(* IEC 61131-3 sources: bevling_machine/framework/sources/04_Machine, 9 files *)

(* ---- F_RecipeValid.st ---- *)
(* 模块说明：检查框架允许的料型、速度、行程和位置顺序。通过仅表示符合示例边界，不代表实机参数已经确认。 *)
FUNCTION F_RecipeValid : BOOL
VAR_INPUT
    stRecipe : ST_Recipe; (* 待校验配方或上层传入的运行配方，字段含义见 ST_Recipe。 *)
END_VAR
FUNCTION F_RecipeValid : BOOL
(* 示例边界：切长 0..1200、速度 0..300、角度正负360，并要求机械手回位<后退<前进<拉料。边界是否适合实机仍需标定。 *)
(* 料型只认 300/450/600：现场侧挡是三个固定位置的气缸，没有 400 这个档；400 是早期仿真的占位值。 *)
F_RecipeValid := ((stRecipe.uiMaterialModel = 300) OR
    (stRecipe.uiMaterialModel = 450) OR (stRecipe.uiMaterialModel = 600))
    AND (stRecipe.lrCutLength > 0.0) AND (stRecipe.lrCutLength <= 1200.0)
    AND (stRecipe.lrCutVelocity > 0.0) AND (stRecipe.lrCutVelocity <= 300.0)
    AND (stRecipe.lrReturnVelocity > 0.0) AND (stRecipe.lrReturnVelocity <= 300.0)
    AND (stRecipe.lrPositionVelocity > 0.0) AND (stRecipe.lrPositionVelocity <= 100.0)
    AND (stRecipe.lrBeltVelocity > 0.0) AND (stRecipe.lrBeltVelocity <= 100.0)
    AND (stRecipe.lrSpindleVelocity > 0.0) AND (stRecipe.lrSpindleVelocity <= 100.0)
    AND (stRecipe.tStepTimeout >= T#1S) AND (stRecipe.tCutTimeout >= T#1S) AND (stRecipe.tSpray > T#0MS)
    AND (ABS(stRecipe.lrCutHome) <= 500.0)
    (* 终点 = 回刀起点 + 切割行程；行程放到 1200 后，终点上限相应放到 1300（典型 100+1200）。 *)
    AND (ABS(stRecipe.lrCutHome + stRecipe.lrCutLength) <= 1300.0)
    AND (ABS(stRecipe.lrLengthPosition) <= 1000.0)
    AND (ABS(stRecipe.lrLengthClear) <= 1000.0)
    AND (ABS(stRecipe.lrRotateAngle) <= 360.0)
    AND (stRecipe.lrGripperHome < stRecipe.lrGripperBack)
    AND (stRecipe.lrGripperBack < stRecipe.lrGripperFront)
    AND (stRecipe.lrGripperFront < stRecipe.lrGripperPull)
    AND (ABS(stRecipe.lrGripperPull) <= 1000.0);

(* ---- FB_AlarmManager.st ---- *)
(* 模块说明：锁存首次非零报警。只有复位有效且当前没有新报警时清除；同一扫描有新报警时仍会锁存。 *)
FUNCTION_BLOCK FB_AlarmManager
VAR_INPUT
    udiIncoming : UDINT; (* 当前扫描的新报警码；0 表示当前未提出报警。 *)
    xReset : BOOL; (* 故障复位许可；仿真设备仅在故障注入已撤销时清除错误。 *)
END_VAR
VAR_OUTPUT
    udiLatched : UDINT; (* 已锁存的首个非零报警码；后续报警不覆盖，满足复位条件后清零。 *)
END_VAR
FUNCTION_BLOCK FB_AlarmManager
(* 只有没有当前报警原因才清锁存；当前代码保留第一个非零报警，后续报警不覆盖。 *)
IF xReset AND (udiIncoming=0) THEN udiLatched:=0; END_IF
IF (udiLatched=0) AND (udiIncoming<>0) THEN udiLatched:=udiIncoming; END_IF

(* ---- FB_AutoCycle.st ---- *)
(* 模块说明：自动主状态机。只组织工序并提出请求，设备执行由整机统一调用；送料等料允许长期等待。 *)
FUNCTION_BLOCK FB_AutoCycle
VAR_INPUT
    xRun : BOOL; (* 自动工序运行许可，整机 Automatic 时保持 TRUE；撤销立即复位主流程。 *)
    xContinuous : BOOL; (* TRUE 连续循环；FALSE 在当前完整循环结束后回到就绪。 *)
    xMaterialAtLength : BOOL; (* 定长光电到位状态；自动送料须先离开再到位，并满足 D5 下降。 *)
    stRecipe : ST_Recipe; (* 待校验配方或上层传入的运行配方，字段含义见 ST_Recipe。 *)
END_VAR
VAR_IN_OUT
    aCommand : ARRAY[1..17] OF ST_DeviceCommand; (* 统一设备请求数组 1..17；子流程写请求，设备管理器执行。 *)
    aStatus : ARRAY[1..17] OF ST_DeviceStatus; (* 各设备的反馈数组 1..17，供判断忙、完成序号、故障和位置。 *)
    udiCounter : UDINT; (* 全机共享的动作序号计数器，通过引用传递；由 F_NextID 分配，0 不使用。 *)
END_VAR
VAR_OUTPUT
    eStep : E_AutoStep; (* 自动主工序当前状态，见 E_AutoStep。 *)
    xDone : BOOL; (* 整循环完成的单扫描脉冲；机械手等三路收尾全部结束后才产生。 *)
    xError : BOOL; (* 本设备或本子流程发生故障；具体原因见对应错误码。 *)
    udiErrorID : UDINT; (* 非法主步骤为 4800；主步超时为 4800+步号；步骤守护失败为 4800+步号+1，见下方守护表；支线错误则向上传递。 *)
    uiClearLengthStep : UINT; (* 避让支线 P 的当前步骤：10 升起 D5，20 移开 D4，1000 完成。 *)
    uiClearTransferStep : UINT; (* 避让支线 Q 当前步骤：10 降 G4，20 松 G3，30 降 G2，1000 完成。 *)
    uiPostStep : UINT; (* 收尾总步骤：10 抬刀，20 抬压，30 等待三路完成，1000 结束。 *)
    uiReturnKnifeStep : UINT; (* 收尾支线 A：10 喷油，20 D2 回刀，1000 完成。 *)
    uiUnloadStep : UINT; (* 机械手移料支线 B 步骤，10..110 每步加 10，1000 完成；详见 FB_Unload。 *)
    uiResetLengthStep : UINT; (* 收尾支线 C：10 D4 定位，20 D5 下降，30 确认下降，1000 完成。 *)
END_VAR
VAR
    ePrevStep : E_AutoStep := E_AutoStep.Fault; (* 上扫描主工序状态，用于产生步骤入口标志。 *)
    udiToken : UDINT; (* 本步骤专用动作序号；同一步中的设备共用该号，以排除旧完成信号。 *)
    udiSpindleToken : UDINT; (* 盘刀运行命令序号，切割过程中保持该号，避免重复重启盘刀命令。 *)
    udiPressToken : UDINT; (* G1 下压保位序号；PressDown 入口分配，后续步骤持续用该号重发，保证单电控阀不断电。 *)
    udiKnifeToken : UDINT; (* G9 下刀保位序号；KnifeDown 入口分配，同上。 *)
    xEntry : BOOL; (* 本扫描为新步骤入口；用于分配新序号并复位步骤超时计时。 *)
    xSawSensorClear : BOOL; (* 本轮送料已观察到光电离开；须先有该标志再接受新到位，防止残留信号触发。 *)
    tonStep : TON; (* 步骤超时定时器；进入新步骤时复位，超时错误码由模块及当前步号组成。 *)
    tStepLimit : TIME; (* 本扫描用的步骤超时值：切割步取 tCutTimeout，其余取 tStepTimeout。 *)
    xGuardOK : BOOL; (* 步骤守护判据：当前步依赖的前提是否仍满足，FALSE 时立即报错退出，不等步超时。 *)
    fbClear : FB_ClearanceUnit; (* 切割前两路并行避让流程。 *)
    fbPost : FB_PostCut; (* 切割后抬刀、抬压及三路收尾流程。 *)
END_VAR
FUNCTION_BLOCK FB_AutoCycle
(* 完成标志每扫描先清零；本流程在许可撤销后复位，不保留中断点续跑。 *)
xDone := FALSE;
IF NOT xRun THEN eStep:=E_AutoStep.Idle; xError:=FALSE; udiErrorID:=0; xSawSensorClear:=FALSE; END_IF
(* 进入新步骤才换新动作序号，同一步持续保持请求，防止反复启动。 *)
xEntry := eStep <> ePrevStep;
IF xEntry THEN udiToken := F_NextID(udiCounter); END_IF
ePrevStep := eStep;
(* 送料等料不计步骤超时；其余执行步按运行配方监控。
   切割步单独用 tCutTimeout：走刀行程长，和其它单动作步共用一个 30 秒很容易误超时。 *)
tStepLimit := stRecipe.tStepTimeout;
IF eStep = E_AutoStep.Cutting THEN tStepLimit := stRecipe.tCutTimeout; END_IF
tonStep(IN:=xRun AND NOT xEntry AND (eStep<>E_AutoStep.Idle)
    AND (eStep<>E_AutoStep.FeedWait) AND (eStep<>E_AutoStep.Complete)
    AND (eStep<>E_AutoStep.Fault),PT:=tStepLimit);
IF xRun AND NOT xError THEN
CASE eStep OF
(* 待机转入送料；没有直接跳到切割。 *)
E_AutoStep.Idle: eStep:=E_AutoStep.FeedWait;
(* D1 送料并正常等料；光电须先离开再到位，且 D5 必须在下降端。 *)
E_AutoStep.FeedWait:
    IF xEntry THEN xSawSensorClear:=FALSE; END_IF
    IF NOT xMaterialAtLength THEN xSawSensorClear:=TRUE; END_IF
    aCommand[1]:=F_Command(E_DeviceAction.Run,udiToken,0.0,stRecipe.lrBeltVelocity);
    IF xSawSensorClear AND xMaterialAtLength AND F_At(aStatus[5],1.0) THEN eStep:=E_AutoStep.StopFeed; END_IF
(* 本步不再给 D1 运行请求，整机周期清空请求后等待皮带非运行、非忙。 *)
E_AutoStep.StopFeed:
    IF NOT aStatus[1].xActive AND NOT aStatus[1].xBusy THEN eStep:=E_AutoStep.Push; END_IF
(* G3 侧推到位；只认本次 udiToken 对应的完成。 *)
E_AutoStep.Push:
    aCommand[11]:=F_Command(E_DeviceAction.Position,udiToken,1.0,stRecipe.lrPositionVelocity);
    IF F_Done(aStatus[11],udiToken) THEN eStep:=E_AutoStep.Clearance; END_IF
(* 并行调用定长避让 P 和输送机构避让 Q，两路都完成后旋转平台。 *)
E_AutoStep.Clearance:
    IF fbClear.xDone THEN eStep:=E_AutoStep.Rotate; END_IF
(* D8 旋转到 lrRotateAngle，必须在 G1 下压之前完成。 *)
E_AutoStep.Rotate:
    aCommand[8]:=F_Command(E_DeviceAction.Position,udiToken,stRecipe.lrRotateAngle,stRecipe.lrPositionVelocity);
    IF F_Done(aStatus[8],udiToken) THEN eStep:=E_AutoStep.PressDown; END_IF
(* G1 下压到位。 *)
E_AutoStep.PressDown:
    IF xEntry THEN udiPressToken:=udiToken; END_IF
    aCommand[9]:=F_Command(E_DeviceAction.Position,udiPressToken,1.0,stRecipe.lrPositionVelocity);
    IF F_Done(aStatus[9],udiPressToken) THEN eStep:=E_AutoStep.SpindleOn; END_IF
(* D3 盘刀先转起来，转稳了再下刀；此时刀还没下来，G1 保持压紧。 *)
E_AutoStep.SpindleOn:
    udiSpindleToken:=udiToken;
    aCommand[9]:=F_Command(E_DeviceAction.Position,udiPressToken,1.0,stRecipe.lrPositionVelocity);
    aCommand[3]:=F_Command(E_DeviceAction.Run,udiSpindleToken,0.0,stRecipe.lrSpindleVelocity);
    IF F_Done(aStatus[3],udiSpindleToken) AND aStatus[3].xActive THEN eStep:=E_AutoStep.KnifeDown; END_IF
(* G9 盘刀下降到位；下降全程 D3 保持运行。 *)
E_AutoStep.KnifeDown:
    IF xEntry THEN udiKnifeToken:=udiToken; END_IF
    aCommand[9]:=F_Command(E_DeviceAction.Position,udiPressToken,1.0,stRecipe.lrPositionVelocity);
    aCommand[3]:=F_Command(E_DeviceAction.Run,udiSpindleToken,0.0,stRecipe.lrSpindleVelocity);
    aCommand[17]:=F_Command(E_DeviceAction.Position,udiKnifeToken,1.0,stRecipe.lrPositionVelocity);
    IF F_Done(aStatus[17],udiKnifeToken) THEN eStep:=E_AutoStep.Cutting; END_IF
(* 保持 D3 运行，G6 吹气，D2 走到回刀起点加切割长度；以 D2 到位作为切割完成。 *)
E_AutoStep.Cutting:
    aCommand[9]:=F_Command(E_DeviceAction.Position,udiPressToken,1.0,stRecipe.lrPositionVelocity);
    aCommand[17]:=F_Command(E_DeviceAction.Position,udiKnifeToken,1.0,stRecipe.lrPositionVelocity);
    aCommand[3]:=F_Command(E_DeviceAction.Run,udiSpindleToken,0.0,stRecipe.lrSpindleVelocity);
    aCommand[14]:=F_Command(E_DeviceAction.Run,udiToken,0.0,0.0);
    aCommand[2]:=F_Command(E_DeviceAction.Position,udiToken,stRecipe.lrCutHome+stRecipe.lrCutLength,stRecipe.lrCutVelocity);
    IF F_Done(aStatus[2],udiToken) THEN eStep:=E_AutoStep.StopCut; END_IF
(* 撤销 D3/G6 运行请求，等待盘刀停止且吹气关闭后收尾。 *)
E_AutoStep.StopCut:
    aCommand[9]:=F_Command(E_DeviceAction.Position,udiPressToken,1.0,stRecipe.lrPositionVelocity);
    aCommand[17]:=F_Command(E_DeviceAction.Position,udiKnifeToken,1.0,stRecipe.lrPositionVelocity);
    IF NOT aStatus[3].xActive AND NOT aStatus[3].xBusy AND NOT aStatus[14].xActive THEN eStep:=E_AutoStep.PostCut; END_IF
(* 先抬刀再抬压，随后三支线同步执行；全部结束才完成本轮。 *)
E_AutoStep.PostCut:
    IF fbPost.xDone THEN eStep:=E_AutoStep.Complete; END_IF
(* 只在进入本步时输出一次完成脉冲；连续模式返回送料，单循环由整机回到 Ready。 *)
E_AutoStep.Complete:
    xDone:=xEntry;
    IF xContinuous THEN eStep:=E_AutoStep.FeedWait; END_IF
(* 保留流程错误状态；整机退出自动后才复位此流程。 *)
E_AutoStep.Fault: xError:=TRUE;
ELSE xError:=TRUE; udiErrorID:=4800;
END_CASE
(* ===== 步骤守护表 =====
   只判前提，不判目标：目标是本步自己要去达成的东西，由各步的 F_Done 判完成；
   这里判的是这一步所依赖的前提还在不在。前提在进入该步时就已成立，
   之后必须一直保持，一旦丢失立即报错退出，不再干等 tonStep 超时才发现。
   每个步骤都要在下面有明确交代，无守护也要写出来，避免以后分不清
   是真的不需要还是漏掉了。新增步骤时先到这里补一行。
   错误码约定：4800 + 步号 + 1，例 SpindleOn=4881、Cutting=4891。
   这里不主动发 Stop：报错后本流程转 Fault，下一扫描不再提出任何请求，
   设备管理器收到 None 即停止，轴走 MC_Stop，气缸阀失电。 *)
xGuardOK := TRUE;
CASE eStep OF
(* 无守护：要么在等外部条件，要么本步本身就在建立条件。 *)
E_AutoStep.Idle, E_AutoStep.FeedWait, E_AutoStep.StopFeed,
E_AutoStep.Push, E_AutoStep.Clearance, E_AutoStep.Rotate,
E_AutoStep.PressDown, E_AutoStep.StopCut,
E_AutoStep.PostCut, E_AutoStep.Complete, E_AutoStep.Fault:
    xGuardOK := TRUE;

(* 起盘刀前：只要已压紧；此时刀还没下来，不判下刀。 *)
E_AutoStep.SpindleOn:
    xGuardOK := F_At(aStatus[9],1.0);

(* 下刀期间：压紧且盘刀必须已经在转，不能拿一把没转的刀往下扎。 *)
E_AutoStep.KnifeDown:
    xGuardOK := F_At(aStatus[9],1.0) AND aStatus[3].xActive;

(* 切割全程：压紧、下刀、盘刀运行三者都必须保持。 *)
E_AutoStep.Cutting:
    xGuardOK := F_At(aStatus[9],1.0) AND F_At(aStatus[17],1.0) AND aStatus[3].xActive;
END_CASE
IF NOT xGuardOK THEN
    xError := TRUE;
    udiErrorID := 4800 + TO_UDINT(eStep) + 1;
END_IF
IF tonStep.Q THEN xError:=TRUE; udiErrorID:=4800+TO_UDINT(eStep); END_IF
END_IF
(* 子功能块必须每扫描调用，包括失能时复位；上方状态判断看到的是此前反馈。 *)
fbClear(xExecute:=xRun AND (eStep=E_AutoStep.Clearance),stRecipe:=stRecipe,aCommand:=aCommand,aStatus:=aStatus,udiCounter:=udiCounter);
fbPost(xExecute:=xRun AND (eStep=E_AutoStep.PostCut),stRecipe:=stRecipe,aCommand:=aCommand,aStatus:=aStatus,udiCounter:=udiCounter);
(* 任一支线错误向主流程上报；所有设备请求还须经过整机统一互锁。 *)
IF fbClear.xError OR fbPost.xError THEN xError:=TRUE; udiErrorID:=MAX(fbClear.udiErrorID,fbPost.udiErrorID); END_IF
IF xError THEN eStep:=E_AutoStep.Fault; END_IF
uiClearLengthStep:=fbClear.uiLengthStep; uiClearTransferStep:=fbClear.uiTransferStep;
uiPostStep:=fbPost.uiStep; uiReturnKnifeStep:=fbPost.uiKnifeStep;
uiUnloadStep:=fbPost.uiUnloadStep; uiResetLengthStep:=fbPost.uiLengthStep;

(* ---- FB_Indicator.st ---- *)
(* 模块说明：面板两色指示灯的纯输出逻辑。指示灯没有反馈、不参与互锁、不占设备索引，
   所以不做成设备，只在这里按整机状态算出两个灯的电平，由 PLC_PRG 下沉到 GVL_IO_Physical。
   优先级：停止/故障最高（红亮绿灭）→ 自动循环运行中（绿慢闪）→ 其余正常运行（绿常亮）。 *)
FUNCTION_BLOCK FB_Indicator
VAR_INPUT
	xRunState : BOOL; (* 整机运行态锁存；FALSE 表示按过停止或上电还没启动。 *)
	eState : E_MachineState; (* 整机状态；Stopped 与 Fault 一律按停机处理。 *)
	eMode : E_MachineMode; (* 模式旋钮当前选择；只有自动循环真正在跑时绿灯才改为慢闪。 *)
	udiAlarm : UDINT; (* 锁存报警码；非 0 时按故障处理，红亮绿灭。 *)
	tBlinkHalf : TIME := T#500MS; (* 慢闪半周期：500 ms 亮 + 500 ms 灭，即每秒亮灭一次。 *)
END_VAR
VAR_OUTPUT
	xGreen : BOOL; (* 绿灯电气电平，TRUE 为亮。 *)
	xRed : BOOL; (* 红灯电气电平，TRUE 为亮。 *)
	xBlinking : BOOL; (* 绿灯当前处于闪烁状态；仅用于监控，不参与控制。 *)
END_VAR
VAR
	tonBlink : TON; (* 闪烁节拍定时器；到点翻转相位并自复位，形成连续方波。 *)
	xBlinkPhase : BOOL; (* 闪烁相位：TRUE 为亮的那一半。 *)
END_VAR
FUNCTION_BLOCK FB_Indicator
(* 先算闪烁节拍：定时器到点就翻转相位并自复位，得到占空比 50% 的连续方波。
   IN 取 Q 的反相做自复位，Q 每次只保持一个扫描，正好当翻转脉冲用。 *)
tonBlink(IN := NOT tonBlink.Q, PT := tBlinkHalf);
IF tonBlink.Q THEN xBlinkPhase := NOT xBlinkPhase; END_IF

(* 停机判据与状态机保持同一口径：运行态锁存为假、处在故障、或有锁存报警，都算停下。
   红灯优先，任何情况下都不会出现红绿同时亮。 *)
IF (NOT xRunState) OR (eState = E_MachineState.Fault) OR (udiAlarm <> 0) THEN
	xRed := TRUE; xGreen := FALSE; xBlinking := FALSE;
(* 自动循环运行中：绿灯慢闪，表示"正在自动动作"，与手动时有人在场操作区分开。 *)
ELSIF (eMode = E_MachineMode.Automatic) AND (eState = E_MachineState.Automatic) THEN
	xRed := FALSE; xGreen := xBlinkPhase; xBlinking := TRUE;
(* 其余运行状态（手动、初始化中、已就绪待启动）：绿灯常亮。 *)
ELSE
	xRed := FALSE; xGreen := TRUE; xBlinking := FALSE;
END_IF

(* ---- FB_Interlocks.st ---- *)
(* 模块说明：对手动、初始化和自动请求统一执行软件互锁。禁止动作时改为停止，并报告最后一个被阻挡设备。 *)
FUNCTION_BLOCK FB_Interlocks
VAR_INPUT
	xPermit : BOOL; (* 整机当前允许发出动作的总许可；仍需继续满足各设备互锁。 *)
	xManualMode : BOOL; (* 当前处于手动模式；手动模式暂不做机构互锁，互锁只约束自动流程。 *)
	stRecipe : ST_Recipe; (* 待校验配方或上层传入的运行配方，字段含义见 ST_Recipe。 *)
	stReal : ST_RealDeviceSettings; (* 真实设备接管设置；预留输入，当前手动已默认不查互锁，判定未使用。 *)
    tViolationDelay : TIME := T#200MS; (* 机构违规确认时间；连续保持这么久才认定，避免过渡瞬间误报。 *)
	aRequest : ARRAY[1..17] OF ST_DeviceCommand; (* 初始化/手动/自动产生的原始请求，每周期先清空，再交互锁筛选。 *)
	aStatus : ARRAY[1..17] OF ST_DeviceStatus; (* 各设备的反馈数组 1..17，供判断忙、完成序号、故障和位置。 *)
END_VAR
VAR_OUTPUT
	aCommand : ARRAY[1..17] OF ST_DeviceCommand; (* 统一设备请求数组 1..17；子流程写请求，设备管理器执行。 *)
	uiBlockedDevice : UINT; (* 本扫描最后一个被互锁阻挡的设备索引；0 表示无阻挡，可结合设备状态排查。 *)
    xViolated : BOOL; (* 机构互锁违规已确认：总许可通过、但机构条件不满足，且持续超过确认时间。 *)
    uiViolatedDevice : UINT; (* 确认违规的设备索引；0 表示无。 *)
END_VAR
VAR
	i : INT; (* 本扫描数组遍历索引；含义及范围以当前 FOR 循环为准。 *)
	xAllowed : BOOL; (* 当前遍历设备的最终互锁允许结果。 *)
	xMotion : BOOL; (* 当前请求是否为点动或离开当前位置的定位，决定是否检查机构避让。 *)
	xKnifeUp : BOOL; (* G9 刀具处于提升端且设备无忙无故障。 *)
	xPressUp : BOOL; (* G1 下压机构处于抬起端且设备无忙无故障。 *)
	xClampOpen : BOOL; (* G8 夹爪处于打开端且设备无忙无故障。 *)
    xPermitOK : BOOL; (* 仅总许可结果；用来区分"许可没通过"和"机构条件不满足"。 *)
    xStructBlocked : BOOL; (* 本扫描是否有请求因机构条件被拒。 *)
    uiStructDevice : UINT; (* 最后一个因机构条件被拒的设备索引。 *)
    tonViolation : TON; (* 机构违规去抖定时器。 *)
END_VAR
FUNCTION_BLOCK FB_Interlocks
(* 以下为普通程序互锁；实际急停、门锁、失气等安全功能须由最终硬件方案实现。 *)
uiBlockedDevice:=0;
    xStructBlocked:=FALSE;
    uiStructDevice:=UINT#0;
xKnifeUp:=F_At(aStatus[17],0.0); xPressUp:=F_At(aStatus[9],0.0);
xClampOpen:=F_At(aStatus[16],0.0);
FOR i:=1 TO 17 DO
    aCommand[i]:=aRequest[i];
    xPermitOK:=xPermit AND (i<>6);
    xAllowed:=xPermitOK;
    xMotion:=(aRequest[i].eAction=E_DeviceAction.Jog) OR
        ((aRequest[i].eAction=E_DeviceAction.Position) AND
        (ABS(aRequest[i].lrTarget-aStatus[i].lrPosition)>0.01));
    (* 手动模式暂不做机构互锁：单轴调试要求能独立动作，互锁只约束自动流程。
       手动下的硬干涉（D5 挡 D4 行程、平台旋转扫刀等）后续按调试情况逐条补回。
       xPermit 不受此影响，任何时候都要先满足。 *)
    IF xMotion AND NOT xManualMode THEN
        CASE i OF
        (* D4 平移之前，D5 定长升降必须已经升起。 *)
        4: xAllowed:=xAllowed AND F_At(aStatus[5],0.0);
        (* D8 平台旋转之前，盘刀和下压抬起、G3 侧推解除。 *)
        8: xAllowed:=xAllowed AND xKnifeUp AND xPressUp AND F_At(aStatus[11],0.0);
        (* G1 下压时，平台不得旋转，盘刀抬起且 D2 在回刀起点。 *)
        9:
            IF aRequest[i].lrTarget>0.5 THEN
                xAllowed:=xAllowed AND NOT aStatus[8].xBusy AND xKnifeUp AND F_At(aStatus[2],stRecipe.lrCutHome);
            ELSE
                (* 抬起前盘刀必须先抬起，否则刀还在工件里就松了压板。 *)
                xAllowed:=xAllowed AND xKnifeUp;
            END_IF
        (* G9 下刀时，下压到位、旋转停止、定长升起、流利条下降、侧挡下降。 *)
        17:
            IF aRequest[i].lrTarget>0.5 THEN
                xAllowed:=xAllowed AND F_At(aStatus[9],1.0) AND NOT aStatus[8].xBusy
                    AND F_At(aStatus[5],0.0) AND F_At(aStatus[12],0.0) AND F_At(aStatus[10],1.0);
            END_IF
        (* D2 正向切割需下压和盘刀下降到位且盘刀运行；回刀需盘刀抬起。 *)
        2:
            IF ((aRequest[i].eAction=E_DeviceAction.Position) AND (aRequest[i].lrTarget>stRecipe.lrCutHome+0.01))
               OR ((aRequest[i].eAction=E_DeviceAction.Jog) AND (aRequest[i].lrVelocity>0.0)) THEN
                xAllowed:=xAllowed AND F_At(aStatus[9],1.0) AND F_At(aStatus[17],1.0) AND aStatus[3].xActive;
            ELSE xAllowed:=xAllowed AND xKnifeUp;
            END_IF
        (* D7 机械手分点动、拉料、抬升平移与下降回位分别校验，保持后退/下降/回位顺序。 *)
        7:
            xAllowed:=xAllowed AND xKnifeUp AND xPressUp;
            IF aRequest[i].eAction=E_DeviceAction.Jog THEN
                xAllowed:=xAllowed AND F_At(aStatus[15],1.0) AND xClampOpen;
            ELSIF ABS(aRequest[i].lrTarget-stRecipe.lrGripperHome)<0.01 THEN
                xAllowed:=xAllowed AND F_At(aStatus[15],0.0) AND xClampOpen;
            ELSIF ABS(aRequest[i].lrTarget-stRecipe.lrGripperPull)<0.01 THEN
                xAllowed:=xAllowed AND F_At(aStatus[15],1.0) AND F_At(aStatus[16],1.0);
            ELSE xAllowed:=xAllowed AND F_At(aStatus[15],1.0) AND xClampOpen;
            END_IF
        END_CASE
    END_IF
    (* 互锁不满足则用 Stop 覆盖该设备请求；记录最后一个被阻挡编号，便于排查。 *)
    IF NOT xAllowed THEN
        IF aRequest[i].eAction<>E_DeviceAction.None THEN
            uiBlockedDevice:=INT_TO_UINT(i);
            (* 只有总许可通过时的拒绝才算机构违规；许可未通过已由 1001 等上报，不在这里重复。 *)
            IF xPermitOK THEN
                xStructBlocked:=TRUE;
                uiStructDevice:=INT_TO_UINT(i);
            END_IF
        END_IF
        aCommand[i].eAction:=E_DeviceAction.Stop;
    END_IF
END_FOR
tonViolation(IN:=xStructBlocked,PT:=tViolationDelay);
xViolated:=tonViolation.Q;
IF xViolated THEN uiViolatedDevice:=uiStructDevice; ELSE uiViolatedDevice:=UINT#0; END_IF

(* ---- FB_IOMap.st ---- *)
FUNCTION_BLOCK FB_IOMap
(* 模块说明：设备输出到物理 I/O 的唯一下沉点。真实气缸的阀电平在此写到 GVL_IO_Physical，
   同时仍维护逻辑输出数组供诊断观察。G2 三个侧挡阀在这里按料型逐路下沉。 *)
VAR_INPUT
    aCommand : ARRAY[1..17] OF ST_DeviceCommand; (* 最终设备命令，当前仅用于诊断，不直接驱动输出。 *)
    aStatus : ARRAY[1..17] OF ST_DeviceStatus; (* 各设备的反馈数组 1..17，供判断忙、完成序号、故障和位置。 *)
    aValveOut : ARRAY[1..17] OF BOOL; (* 设备管理器给出的阀电气电平 1..17，真实气缸在此下沉到物理点。 *)
    aValveOutAux : ARRAY[1..17] OF BOOL; (* 第二个执行器的阀电气电平 1..17；G1 右压板在此下沉到物理点。 *)
    aG2Valve : ARRAY[1..3] OF BOOL; (* G2 三个侧挡阀电气电平 1=300，2=450，3=600。 *)
    uiG2Band : UINT; (* G2 当前实际下降的料型带号 300/450/600；0 表示三缸全部提升。 *)
END_VAR
VAR_IN_OUT
    axOutputs : ARRAY[0..31] OF BOOL; (* 逻辑数字输出数组 0..31，按阀电平填写，供在线监视与后续扩展。 *)
END_VAR
VAR
    i : INT; (* 本扫描数组遍历索引；含义及范围以当前 FOR 循环为准。 *)
END_VAR
FUNCTION_BLOCK FB_IOMap
(* 逻辑输出先清零，只由下面明确赋值的位置置位；未被接管的气缸输出保持失电。 *)
FOR i:=0 TO 31 DO axOutputs[i]:=FALSE; END_FOR

(* ===== 1. 真实气缸阀输出：直接写物理映射符号，TRUE=阀得电=设备动作 ===== *)
(* 未接管时 aValveOut / aG2Valve 为 FALSE，物理点随之失电，不会带着上一个状态一直通电。 *)
GVL_IO_Physical.xDoG1ValveL := aValveOut[9];
GVL_IO_Physical.xDoG1ValveR := aValveOutAux[9];
GVL_IO_Physical.xDoG2Valve300 := aG2Valve[1];
GVL_IO_Physical.xDoG2Valve450 := aG2Valve[2];
GVL_IO_Physical.xDoG2Valve600 := aG2Valve[3];
GVL_IO_Physical.xDoG3Valve := aValveOut[11];
GVL_IO_Physical.xDoG9Valve := aValveOut[17];

(* ===== 2. G2 当前料型带号：供诊断观察，不再从下降反馈反推 ===== *)
GVL_IO.uiG2BandActive := uiG2Band;

(* ===== 3. 逻辑输出镜像：便于在监视表按索引观察，不直接对应物理点 ===== *)
axOutputs[0] := aValveOut[9];
axOutputs[1] := aG2Valve[1];
axOutputs[2] := aG2Valve[2];
axOutputs[3] := aG2Valve[3];
axOutputs[4] := aValveOut[11];
axOutputs[5] := aValveOut[17];

(* ---- FB_Machine.st ---- *)
(* 模块说明：整机调度中心：命令选择、模式和报警管理、初始化/手动/自动调度、统一互锁、设备执行及状态发布。 *)
FUNCTION_BLOCK FB_Machine
VAR_INPUT
	xSimulation : BOOL; (* TRUE 使用内部仿真；当前 FALSE 报未实现 3001，不会接管真实运动。 *)
	stPanel : ST_OperatorCommand; (* 本地实体面板解码结果；模式、初始化、复位始终以它为准。 *)
	stRemote : ST_RemoteCommand; (* 上位机可选的启停请求，不包含模式或初始化/复位字段。 *)
	xRemoteRequest : BOOL; (* 远程新命令有效脉冲；无新帧时仅保留模式与连续选择。 *)
	xAllowRemoteStartStop : BOOL; (* 本地工程配置授权远程启停，默认 FALSE；不授予改模式、初始化或复位权限，也不映射给上位机写。 *)
	wRemoteSequence : WORD; (* 本次远程新命令序号，整机处理后写入确认状态。 *)
	aManual : ARRAY[1..17] OF ST_ManualCommand; (* 各设备手动请求，索引 1..17；进入手动后先释放所有按钮再允许动作。 *)
	stRecipe : ST_Recipe; (* 待校验配方或上层传入的运行配方，字段含义见 ST_Recipe。 *)
	stSim : ST_SimulationSettings; (* 软件仿真设置；设备管理器按设备索引读取卡住与故障注入。 *)
	stReal : ST_RealDeviceSettings; (* 真实设备接管设置；逐台位决定哪些编号走真实轴。 *)
	xRealSafetyOK : BOOL; (* 真实安全许可预留接口；当前仿真模式使用 stSim.xSafetyOK。 *)
	xRealMaterial : BOOL; (* 真实定长光电预留输入；当前仿真模式由 FB_SimPlant 提供。 *)
	xSafetyBypassActive : BOOL; (* 安全许可两级旁路已生效；仅在 xAnyReal 为 TRUE 时参与取或。 *)
END_VAR
VAR_OUTPUT
	stStatus : ST_MachineStatus; (* 本模块对外发布的状态；字段含义见其数据类型。 *)
	aDeviceStatus : ARRAY[1..17] OF ST_DeviceStatus; (* 设备管理器汇总反馈，索引 1..17；供工序判断及在线监控。 *)
	aSelectedCommand : ARRAY[1..17] OF ST_DeviceCommand; (* 通过统一互锁后的最终设备请求，交设备管理器执行。 *)
	aValveOut : ARRAY[1..17] OF BOOL; (* 各设备阀电气电平，索引同设备号；供物理映射层下沉到真实输出点。 *)
	aValveOutAux : ARRAY[1..17] OF BOOL; (* 第二个执行器的阀电气电平，索引同设备号；当前只有 G1 双压板使用。 *)
	aG2Valve : ARRAY[1..3] OF BOOL; (* G2 三个侧挡阀电气电平 1=300，2=450，3=600；供物理映射层下沉。 *)
	uiG2Band : UINT; (* G2 当前实际下降的料型带号 300/450/600；0 表示三缸全部提升。 *)
END_VAR
VAR
	stCommand : ST_OperatorCommand; (* 本周期选择并合并后的整机命令；本地停止始终优先于远程。 *)
	stActiveRecipe : ST_Recipe; (* 本次初始化/自动启动时采纳的配方快照，运行中不直接跟随参数区变化。 *)
	aRequest : ARRAY[1..17] OF ST_DeviceCommand; (* 初始化/手动/自动产生的原始请求，每周期先清空，再交互锁筛选。 *)
	stEmpty : ST_DeviceCommand; (* 默认全零设备命令，每周期用它清空原始请求，未被重新提出的动作自动取消。 *)
	fbDevices : FB_DeviceManager; (* 统一设备管理器，每周期调用一次，汇总各设备反馈。 *)
	fbManual : FB_ManualControl; (* 手动请求转换功能块，须处于手动并已释放全部按钮才使能。 *)
	fbAuto : FB_AutoCycle; (* 自动主流程功能块，仅在整机 Automatic 状态运行。 *)
	fbInitialize : FB_Initialize; (* 初始化功能块，仅在整机 Initializing 状态执行。 *)
	fbInterlocks : FB_Interlocks; (* 所有模式共用的软件互锁，输出最终允许的请求。 *)
	fbPlant : FB_SimPlant; (* 仿真整机来料模型；当前流程读取其上一扫描的到位反馈。 *)
	fbAlarm : FB_AlarmManager; (* 整机首报警锁存功能块。 *)
	rtInitialize : R_TRIG; (* 初始化按钮上升沿检测。 *)
	rtStart : R_TRIG; (* 自动启动按钮上升沿检测。 *)
	rtReset : R_TRIG; (* 报警复位按钮上升沿检测。 *)
	rtRunStart : R_TRIG; (* 启动按钮上升沿：置运行态锁存。 *)
	rtRunStop : R_TRIG; (* 停止按钮上升沿：清运行态锁存（常闭触点在映射层已取反）。 *)
	xRunState : BOOL; (* 运行态锁存：按一下启动置 TRUE，按一下停止/安全丢失/进故障清 FALSE；全机唯一的"允许动作"判据。 *)
	udiCounter : UDINT; (* 全机共享的动作序号计数器，通过引用传递；由 F_NextID 分配，0 不使用。 *)
	udiFault : UDINT; (* 本扫描整理出的报警原因；设备错误使用 10000+设备索引。 *)
	xSafetyOK : BOOL; (* 安全许可接口或仿真许可，TRUE 允许；不等同于安全级急停回路。 *)
	xMaterial : BOOL; (* 当前实际采用的来料信号，仿真与实机预留输入二选一。 *)
	xInitialized : BOOL; (* 初始化完成标志；停止、运行中切换模式或故障会清除。 *)
	xPermit : BOOL; (* 整机当前允许发出动作的总许可；仍需继续满足各设备互锁。 *)
	xRemoteAccepted : BOOL; (* 本扫描远程命令已获授权，用于回传状态拒绝或配方错误。 *)
	xStartRequest : BOOL; (* 本次启动事件=本地启动按钮上升沿或已接受的远程启动帧；两种事件分别处理以免相互吞掉。 *)
	xResetDevices : BOOL; (* 本扫描设备复位脉冲，需复位上升沿、安全许可和仿真模式均满足。 *)
	xLastSimulation : BOOL := TRUE; (* 上扫描仿真开关；切换模式时清除初始化并停止。 *)
	xManualReleased : BOOL; (* 所有手动按钮都已释放，用于避免带着按住命令进入手动。 *)
	xManualArmed : BOOL; (* 本次进入手动后已观察到全部按钮释放；离开手动即清除。 *)
	eActiveMode : E_MachineMode; (* 当前初始化/运行时采纳的操作模式，用于检测运行中切换模式。 *)
	xAnyReal : BOOL; (* 是否有任意设备由真实轴接管；全 FALSE 时后续分支与改造前逐语句一致。 *)
    udiInterlockFault : UDINT; (* 互锁违规码；互锁在报警汇总之后才调用，故本扫描存入、下扫描并入 udiFault。 *)
	xAllHomed : BOOL; (* 所有已接管的真实轴都已完成回零；未接真实轴时为 TRUE，用于状态发布。 *)
	dwRealMask : DWORD; (* 真实设备接管掩码，第 i 位置位表示设备 i 走真实轴；用 DWORD 是因为索引 17 需要第 16 位，WORD 会溢出丢位。 *)
	dwLastRealMask : DWORD; (* 上扫描接管掩码；变化时清除初始化并回 Stopped。 *)
	xLastRelativeVerify : BOOL; (* 上扫描相对验证开关；切换时清除初始化并回 Stopped。 *)
	uiSafetySource : UINT; (* 安全许可来源：0 仿真源，1 真实源，2 调试旁路。 *)
	uiInitReject : UINT; (* 初始化被拒绝的原因：0 未拒绝；回零已并入初始化流程，当前无拒绝分支，字段预留。 *)
	i : INT; (* 本扫描数组遍历索引；含义及范围以当前 FOR 循环为准。 *)
END_VAR
FUNCTION_BLOCK FB_Machine
(* 零、派生混跑标志：axRealDevice 全 FALSE 时 xAnyReal 为 FALSE，后续所有分支与改造前一致。 *)
xAnyReal:=FALSE; dwRealMask:=0;
FOR i:=1 TO 17 DO
    IF stReal.axRealDevice[i] THEN
        xAnyReal:=TRUE;
        dwRealMask:=dwRealMask OR SHL(DWORD#1,i-1);
    END_IF
END_FOR

(* 一、选择命令来源：本地默认优先；远程须授权，本地停止始终有效。 *)
stCommand:=stPanel;
(* 运行态锁存：按一下切换，不靠按钮保持。停止优先——同扫描两个都按下取停止。
   这是全机唯一的"允许动作"判据；下游不再出现单个按钮电平。 *)
rtRunStart(CLK:=stCommand.xRunStart);
rtRunStop(CLK:=stCommand.xRunStop);
IF rtRunStart.Q THEN xRunState:=TRUE; END_IF
IF rtRunStop.Q OR stCommand.xStop THEN xRunState:=FALSE; END_IF
(* 模式、初始化、复位来自实体面板；远程只可追加经过授权的启停，不能替换整份本地命令。 *)
xRemoteAccepted:=FALSE;
IF xRemoteRequest THEN
    stStatus.wRemoteAckSequence:=wRemoteSequence;
    IF xAllowRemoteStartStop THEN
        IF stRemote.xStop THEN
            stCommand.xStop:=TRUE;
            stStatus.uiRemoteResult:=0; xRemoteAccepted:=TRUE;
        ELSIF stRemote.xStart THEN
            IF (stPanel.eMode=E_MachineMode.Automatic)
               AND (stStatus.eState=E_MachineState.Ready) AND xRunState THEN
                stStatus.uiRemoteResult:=0; xRemoteAccepted:=TRUE;
            ELSE stStatus.uiRemoteResult:=3; END_IF
        ELSE stStatus.uiRemoteResult:=2; END_IF
    ELSE stStatus.uiRemoteResult:=1;
    END_IF
END_IF
(* 二、提取初始化/启动/复位上升沿；采样仿真或真实预留输入。 *)
rtInitialize(CLK:=stCommand.xInitialize);
rtStart(CLK:=stCommand.xStart);
(* 本地启动取按钮上升沿，远程启动取新帧脉冲，分别形成事件；本地停止仍优先。 *)
xStartRequest:=rtStart.Q OR (xRemoteAccepted AND stRemote.xStart AND NOT stRemote.xStop);
rtReset(CLK:=stCommand.xResetAlarm);
(* 混跑时安全源改为真实优先：未接安全回路时靠两级旁路放行，旁路生效不报 1001。 *)
IF xAnyReal THEN
    xSafetyOK:=xRealSafetyOK OR xSafetyBypassActive;
    IF stReal.xUseRealMaterial THEN xMaterial:=xRealMaterial;
    ELSE xMaterial:=fbPlant.xMaterialAtLength; END_IF
ELSIF xSimulation THEN xSafetyOK:=stSim.xSafetyOK; xMaterial:=fbPlant.xMaterialAtLength;
ELSE xSafetyOK:=xRealSafetyOK; xMaterial:=xRealMaterial; END_IF
(* 安全许可丢失立即清运行态：急停或旋钮离开许可位后，恢复必须重新按启动，不能自己回到运行。 *)
IF NOT xSafetyOK THEN xRunState:=FALSE; END_IF
(* 安全来源：0 仿真源，1 真实源，2 调试旁路。 *)
IF NOT xAnyReal THEN uiSafetySource:=0;
ELSIF xSafetyBypassActive AND NOT xRealSafetyOK THEN uiSafetySource:=2;
ELSE uiSafetySource:=1; END_IF
(* 三、整理当前报警原因并清空本扫描请求；未被子流程重新提出的动作自动取消。 *)
udiFault:=0;
IF NOT xSafetyOK THEN udiFault:=1001; END_IF
IF udiInterlockFault<>0 THEN udiFault:=udiInterlockFault; END_IF
IF NOT xSimulation THEN udiFault:=3001; END_IF
(* 仿真开关、接管掩码或验证模式变化，均清除初始化并回 Stopped。 *)
IF (xSimulation<>xLastSimulation) OR (dwRealMask<>dwLastRealMask) OR (stReal.xRelativeVerify<>xLastRelativeVerify) THEN
    stStatus.eState:=E_MachineState.Stopped; xInitialized:=FALSE;
END_IF
xLastSimulation:=xSimulation; dwLastRealMask:=dwRealMask; xLastRelativeVerify:=stReal.xRelativeVerify;
FOR i:=1 TO 17 DO
    IF aDeviceStatus[i].xError THEN udiFault:=10000+INT_TO_UDINT(i); END_IF
    aRequest[i]:=stEmpty;
END_FOR
(* 四、运行中切模式、停止或故障会撤销初始化，不能直接接续上一次工序。 *)
IF (stStatus.eState=E_MachineState.Automatic) OR (stStatus.eState=E_MachineState.Manual) THEN
    IF stCommand.eMode<>eActiveMode THEN stStatus.eState:=E_MachineState.Stopped; xInitialized:=FALSE; END_IF
END_IF
(* 停止是运行态锁存的电平判据：按一下停止后锁存一直为 FALSE，直到再按启动。
   这里用 xRunState 而不是按钮电平，是为了让"停着"和"按钮松开"不再有区别。 *)
IF NOT xRunState THEN
    IF (stStatus.eState<>E_MachineState.Stopped) AND (stStatus.eState<>E_MachineState.Fault) THEN
        stStatus.eState:=E_MachineState.Stopped;
    END_IF
    xInitialized:=FALSE;
END_IF
IF udiFault<>0 THEN stStatus.eState:=E_MachineState.Fault; xInitialized:=FALSE; END_IF
(* 五、复位设备和首报警锁存；必须先撤销故障原因，复位不自动启动。 *)
xResetDevices:=rtReset.Q AND xSafetyOK AND xSimulation;
IF xResetDevices THEN
    (* 复位时先按仍有效的故障注入判断原因，再清设备错误和整机锁存；原因未撤销不能复位。 *)
    udiFault:=0;
    udiInterlockFault:=0;
    FOR i:=1 TO 17 DO IF stSim.axFault[i] THEN udiFault:=10000+INT_TO_UDINT(i); END_IF END_FOR
END_IF
fbAlarm(udiIncoming:=udiFault,xReset:=xResetDevices);
IF (stStatus.eState=E_MachineState.Fault) AND (fbAlarm.udiLatched=0) AND xResetDevices THEN
    stStatus.eState:=E_MachineState.Stopped;
END_IF
IF fbAlarm.udiLatched<>0 THEN stStatus.eState:=E_MachineState.Fault; END_IF
(* 六、仅停止态接受初始化；配方通过检查后取快照。 *)
IF rtInitialize.Q AND xRunState THEN
    (* 真实轴的回零已并入初始化第 25 步，这里不再要求预先打开相对验证。 *)
    IF (stStatus.eState=E_MachineState.Stopped) AND xSimulation AND xSafetyOK AND F_RecipeValid(stRecipe) THEN
        stActiveRecipe:=stRecipe; stStatus.eState:=E_MachineState.Initializing;
        eActiveMode:=stCommand.eMode; xInitialized:=FALSE; uiInitReject:=0;
    ELSE
        (* 当前无拒绝分支：回零并入初始化，uiInitReject 保留字段但不再置位。 *)
        IF xRemoteAccepted THEN stStatus.uiRemoteResult:=3; END_IF
    END_IF
END_IF
(* 七、手动不依赖初始化：停机态只要模式在手动且运行态成立就直接进入，开机后不必先跑初始化。
   自动仍必须先完成初始化到 Ready；按过停止后运行态为假，手动也进不去，必须重新按启动。 *)
IF (stStatus.eState=E_MachineState.Stopped) AND (stCommand.eMode=E_MachineMode.Manual)
   AND xRunState THEN
    stStatus.eState:=E_MachineState.Manual; eActiveMode:=E_MachineMode.Manual;
END_IF
IF stStatus.eState=E_MachineState.Ready THEN
    IF stCommand.eMode=E_MachineMode.Manual THEN
        stStatus.eState:=E_MachineState.Manual; eActiveMode:=E_MachineMode.Manual;
    ELSIF xStartRequest AND xRunState THEN
        IF stReal.xRelativeVerify THEN
            (* 相对验证模式下绝对位置不作生产依据，禁止进自动。 *)
            stStatus.uiRemoteResult:=4;
        ELSIF F_RecipeValid(stRecipe) THEN
            stActiveRecipe:=stRecipe; eActiveMode:=E_MachineMode.Automatic;
            stStatus.eState:=E_MachineState.Automatic;
        ELSIF xRemoteAccepted THEN stStatus.uiRemoteResult:=5;
        END_IF
    END_IF
ELSIF (stStatus.eState=E_MachineState.Manual) AND (stCommand.eMode=E_MachineMode.Automatic) THEN
    stStatus.eState:=E_MachineState.Stopped; xInitialized:=FALSE;
END_IF
IF xStartRequest AND xRemoteAccepted AND (stStatus.eState<>E_MachineState.Automatic)
   AND (stStatus.uiRemoteResult=0) THEN stStatus.uiRemoteResult:=3; END_IF

(* 八、手动进入联锁：观察到一次全部按钮释放后，才开放点动/定位操作。 *)
xManualReleased:=TRUE;
FOR i:=1 TO 17 DO
    IF aManual[i].xJogPositive OR aManual[i].xJogNegative OR aManual[i].xMove OR aManual[i].xRun OR aManual[i].xHome THEN xManualReleased:=FALSE; END_IF
END_FOR
IF stStatus.eState<>E_MachineState.Manual THEN xManualArmed:=FALSE;
ELSIF xManualReleased THEN xManualArmed:=TRUE;
END_IF
(* 九、每扫描调用各模式功能块，失能的流程同时复位；共享请求只由当前模式提出。 *)
fbInitialize(xExecute:=stStatus.eState=E_MachineState.Initializing,stRecipe:=stActiveRecipe,
    aCommand:=aRequest,aStatus:=aDeviceStatus,udiCounter:=udiCounter);
fbManual(xEnable:=(stStatus.eState=E_MachineState.Manual) AND xManualArmed,stReal:=stReal,
    aManual:=aManual,aCommand:=aRequest,aStatus:=aDeviceStatus,udiCounter:=udiCounter);
fbAuto(xRun:=stStatus.eState=E_MachineState.Automatic,xContinuous:=stCommand.xContinuous,
    xMaterialAtLength:=xMaterial,stRecipe:=stActiveRecipe,aCommand:=aRequest,aStatus:=aDeviceStatus,udiCounter:=udiCounter);
(* 十、汇总流程完成和流程错误，单循环完成后回到 Ready。 *)
IF fbInitialize.xDone THEN xInitialized:=TRUE; stStatus.eState:=E_MachineState.Ready; END_IF
IF fbInitialize.xError OR fbAuto.xError THEN
    udiFault:=MAX(fbInitialize.udiErrorID,fbAuto.udiErrorID);
    fbAlarm(udiIncoming:=udiFault,xReset:=FALSE);
    stStatus.eState:=E_MachineState.Fault; xInitialized:=FALSE;
END_IF
IF fbAuto.xDone THEN
    stStatus.udiCycleCount:=stStatus.udiCycleCount+1;
    IF NOT stCommand.xContinuous THEN stStatus.eState:=E_MachineState.Ready; END_IF
END_IF
(* 十一、总许可与机构互锁筛选请求，再调用设备管理器；流程判断使用此前的反馈。 *)
xPermit:=xSimulation AND xSafetyOK AND xRunState AND (fbAlarm.udiLatched=0)
    AND ((stStatus.eState=E_MachineState.Initializing) OR (stStatus.eState=E_MachineState.Manual)
    OR (stStatus.eState=E_MachineState.Automatic));
(* 互锁违规先清后置：违规在下面 fbInterlocks 之后才算出，本扫描存入，下扫描并入 udiFault。 *)
udiInterlockFault:=0;
fbInterlocks(xPermit:=xPermit,xManualMode:=(stStatus.eState=E_MachineState.Manual),
    stRecipe:=stActiveRecipe,stReal:=stReal,aRequest:=aRequest,aStatus:=aDeviceStatus);
aSelectedCommand:=fbInterlocks.aCommand;
IF fbInterlocks.xViolated THEN udiInterlockFault:=5000+UINT_TO_UDINT(fbInterlocks.uiViolatedDevice); END_IF
fbDevices(xEnable:=xSimulation AND xSafetyOK,xSimulation:=xSimulation,xReset:=xResetDevices,
    xFaultHold:=(fbAlarm.udiLatched<>0),stSim:=stSim,stReal:=stReal,
    uiMaterialModel:=stActiveRecipe.uiMaterialModel,aCommand:=aSelectedCommand);
aDeviceStatus:=fbDevices.aStatus;
aValveOut:=fbDevices.aValveOut;
aValveOutAux:=fbDevices.aValveOutAux;
aG2Valve:=fbDevices.aG2Valve;
uiG2Band:=fbDevices.uiG2Band;
fbPlant(xEnable:=xSimulation,stSettings:=stSim,aStatus:=aDeviceStatus);
(* 十二、集中发布状态；机械手/定长/回刀卡在哪一步，可从对应 ui...Step 追踪。 *)
(* 故障一律清运行态：故障原因消失后不会自己恢复运行，必须重新按启动。 *)
IF stStatus.eState=E_MachineState.Fault THEN xRunState:=FALSE; END_IF
stStatus.eMode:=stCommand.eMode; stStatus.eAutoStep:=fbAuto.eStep;
stStatus.xSimulation:=xSimulation; stStatus.xRealBackendAvailable:=xAnyReal;
(* 对外掩码仍是 WORD，索引 17（第 16 位）不进这个字段；看真实接管请用 dwRealMask 内部量。 *)
stStatus.xAnyRealDevice:=xAnyReal; stStatus.wRealDeviceMask:=DWORD_TO_WORD(dwRealMask);
stStatus.xRunState:=xRunState;
stStatus.xRelativeVerify:=stReal.xRelativeVerify;
stStatus.xSafetyBypassed:=xSafetyBypassActive AND xAnyReal;
stStatus.uiSafetySource:=uiSafetySource; stStatus.uiInitReject:=uiInitReject;
stStatus.xRemoteStartStopAllowed:=xAllowRemoteStartStop;
xAllHomed:=TRUE;
FOR i:=1 TO 17 DO
    (* D3 盘刀只做连续旋转、不做回零，不参与“全部真实轴已回零”判定，否则该状态永远为 FALSE。 *)
    IF stReal.axRealDevice[i] AND (i<>3) AND (i<9) AND NOT aDeviceStatus[i].xHomed THEN xAllHomed:=FALSE; END_IF
END_FOR
stStatus.xRealAxesHomed:=xAllHomed;
stStatus.xInitialized:=xInitialized;
stStatus.xReady:=xInitialized AND (stStatus.eState=E_MachineState.Ready);
stStatus.xMaterialAtLength:=xMaterial; stStatus.xCycleComplete:=fbAuto.xDone;
stStatus.udiAlarm:=fbAlarm.udiLatched; stStatus.uiBlockedDevice:=fbInterlocks.uiBlockedDevice;
stStatus.uiManualReject:=fbManual.uiRejectDevice;
stStatus.uiClearLengthStep:=fbAuto.uiClearLengthStep; stStatus.uiClearTransferStep:=fbAuto.uiClearTransferStep;
stStatus.uiPostStep:=fbAuto.uiPostStep; stStatus.uiReturnKnifeStep:=fbAuto.uiReturnKnifeStep;
stStatus.uiUnloadStep:=fbAuto.uiUnloadStep; stStatus.uiResetLengthStep:=fbAuto.uiResetLengthStep;
stStatus.uiInitializeStep:=fbInitialize.uiStep; stStatus.uiActiveMaterialModel:=stActiveRecipe.uiMaterialModel;

(* ---- FB_ManualControl.st ---- *)
(* 模块说明：将手动按钮转为统一设备请求。点动松开即取消；定位与回零请求保持到本次完成；D6 不调度。 *)
FUNCTION_BLOCK FB_ManualControl
VAR_INPUT
	xEnable : BOOL; (* 手动模式且按钮释放联锁已满足时允许；未使能也同步按钮快照。 *)
	stReal : ST_RealDeviceSettings; (* 真实设备接管设置；真实编号的手动速度收紧到验证速度。 *)
	aManual : ARRAY[1..17] OF ST_ManualCommand; (* 各设备手动请求，索引 1..17；进入手动后先释放所有按钮再允许动作。 *)
END_VAR
VAR_IN_OUT
	aCommand : ARRAY[1..17] OF ST_DeviceCommand; (* 统一设备请求数组 1..17；子流程写请求，设备管理器执行。 *)
	aStatus : ARRAY[1..17] OF ST_DeviceStatus; (* 各设备的反馈数组 1..17，供判断忙、完成序号、故障和位置。 *)
	udiCounter : UDINT; (* 全机共享的动作序号计数器，通过引用传递；由 F_NextID 分配，0 不使用。 *)
END_VAR
VAR_OUTPUT
	uiRejectDevice : UINT; (* 本扫描最后一个手动拒绝设备索引；0 无，常见原因是冲突按钮或不支持该动作。 *)
END_VAR
VAR
	aPrev : ARRAY[1..17] OF ST_ManualCommand; (* 上扫描手动按钮快照；即使禁用仍更新，防止按住按钮切模式后被误作新上升沿。 *)
	aPending : ARRAY[1..17] OF ST_DeviceCommand; (* 手动定位或回零的锁存请求，直到本次命令完成；点动或运行优先时清除。 *)
	aRunID : ARRAY[1..17] OF UDINT; (* 各设备按住运行/点动时保持的序号，按钮释放后归零。 *)
	i : INT; (* 本扫描数组遍历索引；含义及范围以当前 FOR 循环为准。 *)
	lrVelocity : LREAL; (* 本扫描限幅后的手动速度，取绝对值限幅 0.1..100；反向点动时变为负值。 *)
	lrVelocityMax : LREAL; (* 本扫描速度上限；真实设备收紧到验证速度，防止全速冲出。 *)
	uiPressed : UINT; (* 本扫描该设备同时按下的手动按钮个数；大于 1 视为冲突并拒绝。 *)
END_VAR
FUNCTION_BLOCK FB_ManualControl
(* 每扫描重新判断按钮冲突；无合法请求的设备由整机统一撤销动作。 *)
uiRejectDevice:=0;
FOR i:=1 TO 17 DO
    IF NOT xEnable THEN
        aPending[i].eAction:=E_DeviceAction.None;
        aRunID[i]:=0;
    ELSIF i<>6 THEN
        (* 先撤销本设备请求，只有命中合法按钮时才在下面重新写入。否则松开点动后，
           上一扫描的 Jog 会一直残留在共享请求数组里，真实轴靠 None/Stop 停止的逻辑永远等不到。 *)
        aCommand[i]:=F_Command(E_DeviceAction.None,0,0.0,0.0);
        (* 真实设备的手动速度上限由 lrManualVelocityMax 决定（默认 200）；实际速度取 aManual[i].lrVelocity 与之较小者。 *)
        lrVelocityMax:=100.0;
        IF stReal.axRealDevice[i] THEN
            (* 新字段在未重新初始化的旧下载里可能为 0；兜底 100，避免手动速度变 0 表现为不动作 *)
            lrVelocityMax:=100.0;
            IF stReal.lrManualVelocityMax>0.1 THEN lrVelocityMax:=LIMIT(0.1,stReal.lrManualVelocityMax,200.0); END_IF
        END_IF
        IF i=8 THEN
            (* D8 平台旋转轴（主轴）手动默认 3、限速 5；请求值超过上限时按默认 3 走，不要直接跳到 5。 *)
            lrVelocityMax:=5.0;
            lrVelocity:=3.0;
            IF ABS(aManual[i].lrVelocity)<=lrVelocityMax THEN
                lrVelocity:=LIMIT(0.1,ABS(aManual[i].lrVelocity),lrVelocityMax);
            END_IF
        ELSE
            lrVelocity:=LIMIT(0.1,ABS(aManual[i].lrVelocity),lrVelocityMax);
        END_IF
        (* 任意两个手动按钮同时按下都算冲突：正反点动、点动与定位/运行/回零、定位与运行/回零、运行与回零。 *)
        uiPressed:=0;
        IF aManual[i].xJogPositive THEN uiPressed:=uiPressed+1; END_IF
        IF aManual[i].xJogNegative THEN uiPressed:=uiPressed+1; END_IF
        IF aManual[i].xMove THEN uiPressed:=uiPressed+1; END_IF
        IF aManual[i].xRun THEN uiPressed:=uiPressed+1; END_IF
        IF aManual[i].xHome THEN uiPressed:=uiPressed+1; END_IF
        IF uiPressed>1 THEN
            uiRejectDevice:=INT_TO_UINT(i); aPending[i].eAction:=E_DeviceAction.None;
        (* 点动电平控制，只支持 D2/D4/D5/D7/D8；速度符号决定方向，松开后不保持点动。 *)
        ELSIF aManual[i].xJogPositive OR aManual[i].xJogNegative THEN
            aPending[i].eAction:=E_DeviceAction.None;
            IF aRunID[i]=0 THEN aRunID[i]:=F_NextID(udiCounter); END_IF
            IF aManual[i].xJogNegative THEN lrVelocity:=-lrVelocity; END_IF
            IF (i=2) OR (i=4) OR (i=5) OR (i=7) OR (i=8) THEN
                aCommand[i]:=F_Command(E_DeviceAction.Jog,aRunID[i],0.0,lrVelocity);
            ELSE uiRejectDevice:=INT_TO_UINT(i);
            END_IF
        (* 连续运行电平控制，仅允许皮带、盘刀、喷油和吹气；盘刀接真实轴后走 FB_RealAxis 的 Run 相位。 *)
        ELSIF aManual[i].xRun THEN
            aPending[i].eAction:=E_DeviceAction.None;
            IF (i=1) OR (i=3) OR (i=13) OR (i=14) THEN
                IF aRunID[i]=0 THEN aRunID[i]:=F_NextID(udiCounter); END_IF
                aCommand[i]:=F_Command(E_DeviceAction.Run,aRunID[i],0.0,lrVelocity);
            ELSE uiRejectDevice:=INT_TO_UINT(i);
            END_IF
        (* 回零：上升沿锁存一次请求，之后每扫描重发直到完成；真实轴 D2/D8，D4 为仿真但保留入口。
           D3 盘刀是连续旋转主轴，只做 Run 不做回零，因此不在本白名单内。
           这里不能像点动那样在分支开头清 aPending —— 回零是保持型动作，清了就只剩一个扫描周期，
           设备刚接收就会被下一扫描的 None 撤销，表现为「下发了但不动」。 *)
        ELSIF aManual[i].xHome THEN
            aRunID[i]:=0;
            IF (i=2) OR (i=4) OR (i=8) THEN
                IF NOT aPrev[i].xHome THEN
                    aPending[i]:=F_Command(E_DeviceAction.Home,F_NextID(udiCounter),0.0,0.0);
                END_IF
                IF aPending[i].eAction<>E_DeviceAction.None THEN
                    aCommand[i]:=aPending[i];
                    IF F_Done(aStatus[i],aPending[i].udiID) THEN aPending[i].eAction:=E_DeviceAction.None; END_IF
                END_IF
            ELSE
                (* 不支持的编号：清掉可能从定位继承来的请求，避免继续执行上一个动作。 *)
                uiRejectDevice:=INT_TO_UINT(i);
                aPending[i].eAction:=E_DeviceAction.None;
            END_IF
        ELSE
            aRunID[i]:=0;
            (* 定位仅在按钮上升沿锁存目标和序号，然后持续等待本次完成。 *)
            IF aManual[i].xMove AND NOT aPrev[i].xMove THEN
                IF (i<>1) AND (i<>3) AND (i<>13) AND (i<>14) THEN
                    aPending[i]:=F_Command(E_DeviceAction.Position,F_NextID(udiCounter),aManual[i].lrTarget,lrVelocity);
                ELSE uiRejectDevice:=INT_TO_UINT(i);
                END_IF
            END_IF
            IF aPending[i].eAction<>E_DeviceAction.None THEN
                aCommand[i]:=aPending[i];
                IF F_Done(aStatus[i],aPending[i].udiID) THEN aPending[i].eAction:=E_DeviceAction.None; END_IF
            END_IF
        END_IF
    END_IF
    (* 禁用时仍同步按钮快照，避免按住定位按钮切入手动后产生虚假的新上升沿。 *)
    aPrev[i]:=aManual[i];
END_FOR

(* ---- FB_PanelInput.st ---- *)
(* 模块说明：每扫描先读取实体面板或仿真面板，形成唯一的本地命令来源。上位机不能修改此处的模式。 *)
FUNCTION_BLOCK FB_PanelInput
VAR_INPUT
    xSimulation : BOOL; (* TRUE 使用内部仿真；当前 FALSE 报未实现 3001，不会接管真实运动。 *)
    stReal : ST_PanelInputs; (* 从物理 I/O 映射得到的标准化面板输入，当前未分配端子地址。 *)
    stSim : ST_PanelInputs; (* 仿真用面板输入，代替尚未连接的实体旋钮和按钮。 *)
    xContinuous : BOOL; (* TRUE 连续循环；FALSE 在当前完整循环结束后回到就绪。 *)
    xUseRealPanel : BOOL := TRUE; (* TRUE 取实体面板 stReal；FALSE 取仿真面板 stSim。与 xSimulation 解耦，后者恒为 TRUE。 *)
END_VAR
VAR_OUTPUT
    stCommand : ST_OperatorCommand; (* 由本地面板生成的命令，模式仅由 xAutoMode 形成。 *)
END_VAR
VAR
    stSelected : ST_PanelInputs; (* 本扫描选中的实体/仿真面板输入快照。 *)
END_VAR
FUNCTION_BLOCK FB_PanelInput
(* 这里只处理已归一化的逻辑信号；端子、常开/常闭和必要的输入滤波在实际 I/O 映射时确定。
   面板来源与 xSimulation 解耦：设备可以全仿真而面板用实物按钮，也可以反过来。 *)
IF xUseRealPanel THEN stSelected:=stReal;
ELSE stSelected:=stSim; END_IF
(* 默认手动，只有本地旋钮明确选择自动才转自动；急停反馈不混入普通停止按钮。 *)
stCommand.eMode:=E_MachineMode.Manual;
IF stSelected.xAutoMode THEN stCommand.eMode:=E_MachineMode.Automatic; END_IF
stCommand.xInitialize:=stSelected.xInitialize;
stCommand.xStart:=stSelected.xStart;
stCommand.xStop:=stSelected.xStop;
stCommand.xResetAlarm:=stSelected.xResetAlarm;
stCommand.xContinuous:=xContinuous;
(* 启动/停止是"按一下切换"的两个独立按钮，这里只做电平搬运；
   沿检测与运行态锁存放在 FB_Machine，保证停机判据全机只有一处。 *)
stCommand.xRunStart:=stSelected.xRunStart;
stCommand.xRunStop:=stSelected.xRunStop;
